(* IEC 61131-3 sources: OpenPlc_Lezioni/FlipFlopSR/build, 2 files *)

(* ---- plc.st ---- *)
TYPE
  LOGLEVEL : (CRITICAL, WARNING, INFO, DEBUG) := INFO;
END_TYPE

FUNCTION_BLOCK LOGGER
  VAR_INPUT
    TRIG : BOOL;
    MSG : STRING;
    LEVEL : LOGLEVEL := INFO;
  END_VAR
  VAR
    TRIG0 : BOOL;
  END_VAR

  IF TRIG AND NOT TRIG0 THEN
  {{
   LogMessage(GetFbVar(LEVEL),(char*)GetFbVar(MSG, .body),GetFbVar(MSG, .len));
  }}
  END_IF;
  TRIG0:=TRIG;
END_FUNCTION_BLOCK

PROGRAM program0
  VAR
    SR0 : SR;
    SR1 : SR;
    S1 : BOOL;
    S2 : BOOL;
    RESET : BOOL;
    LED1 : BOOL;
    LED2 : BOOL;
  END_VAR

  SR0(S1 := S1, R := RESET);
  LED1 := SR0.Q1;
  SR1(S1 := S2, R := RESET);
  LED2 := SR1.Q1;
END_PROGRAM

CONFIGURATION Config0

  RESOURCE Res0 ON PLC
    TASK task0(INTERVAL := T#20ms,PRIORITY := 0);
    PROGRAM instance0 WITH task0 : program0;
  END_RESOURCE
END_CONFIGURATION

(* ---- generated_plc.st ---- *)
PROGRAM program0
  VAR
    SR0 : SR;
    SR1 : SR;
    S1 : BOOL;
    S2 : BOOL;
    RESET : BOOL;
    LED1 : BOOL;
    LED2 : BOOL;
  END_VAR

  SR0(S1 := S1, R := RESET);
  LED1 := SR0.Q1;
  SR1(S1 := S2, R := RESET);
  LED2 := SR1.Q1;
END_PROGRAM

CONFIGURATION Config0

  RESOURCE Res0 ON PLC
    TASK task0(INTERVAL := T#20ms,PRIORITY := 0);
    PROGRAM instance0 WITH task0 : program0;
  END_RESOURCE
END_CONFIGURATION
